FUNCTION_BLOCK FsGet (* Copy a file from the file server into a local file *)
  (* Standard: 61499-2; Description: Uses iso_FscReadFileFromServer() of the CCI ISOBUS driver (ISO 11783-13). \n Client is NmDestin.s16OwnCfHnd, file server is NmDestin.s16Handle (e.g. found with NmGetCfInfo, NAME function 61). \n The connection is opened and closed by the driver. One job at a time: REQ during a job gives ERR with s16Status E_BUSY. \n Every REQ ends with exactly one CNF or ERR. \n Local paths: only below /data/fs/, with a logiBUS file server (manufacturer code 1116) below /data/. Paths with .. are refused. \n The local file is replaced; it is written in blocks by a worker task and removed again if the job fails. *)
  (* Version 1.0, 2026-11-25, Franz Höpfinger, initial API and implementation and/or initial documentation *)
  PACKAGE isobus::fs;
  IMPORT isobus::pgn::ISONETEVENT_T;
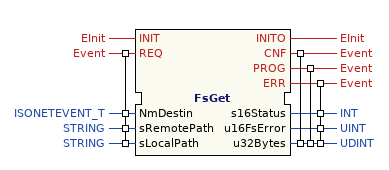
  EVENT_INPUT
    INIT : EInit; (* Service Initialization *)
    REQ WITH NmDestin, sRemotePath, sLocalPath; (* Start the copy *)
  END_EVENT
  EVENT_OUTPUT
    INITO : EInit; (* Initialization Confirm *)
    CNF WITH u32Bytes; (* File copied *)
    PROG WITH u32Bytes; (* Progress (at most every 500 ms) *)
    ERR WITH s16Status, u16FsError, u32Bytes; (* Job failed *)
  END_EVENT
  VAR_INPUT
    NmDestin : isobus::pgn::ISONETEVENT_T; (* Client (s16OwnCfHnd) and file server (s16Handle) *)
    sRemotePath : STRING; (* Path on the file server, e.g. \\USB\data\a.csv *)
    sLocalPath : STRING; (* Local target file, e.g. /data/fs/a.csv *)
  END_VAR
  VAR_OUTPUT
    s16Status : INT; (* With ERR: driver return value or own error (E_BUSY, E_RANGE, E_OVERFLOW) *)
    u16FsError : UINT; (* With ERR: file server or client error (ISO 11783-13 B.9, 6400 ff. client) *)
    u32Bytes : UDINT; (* Bytes copied so far *)
  END_VAR
END_FUNCTION_BLOCK
